Fanuc KAREL source: KD00031.KL

PROGRAM KD00031
%NOLOCKGROUP
VAR
  I: INTEGER
  J: INTEGER
  B: BOOLEAN
  R: REAL
  S: STRING[80]
BEGIN
  CONDITION[1]:
  WHEN PAUSE DO
    I = 1
  ENDCONDITION
END KD00031
